TYPE "FRK_Document_D002"
VERSION : 0.1
   STRUCT
      SchemaVersion { ExternalAccessible := 'False'; ExternalVisible := 'False'; ExternalWritable := 'False'} : UInt;
      Scope { ExternalAccessible := 'False'; ExternalVisible := 'False'; ExternalWritable := 'False'} : String[80];
      Kind { ExternalAccessible := 'False'; ExternalVisible := 'False'; ExternalWritable := 'False'} : DInt;
      ModelCode { ExternalAccessible := 'False'; ExternalVisible := 'False'; ExternalWritable := 'False'} : String[64];
      ActiveModel { ExternalAccessible := 'False'; ExternalVisible := 'False'; ExternalWritable := 'False'} : String[64];
      Count { ExternalAccessible := 'False'; ExternalVisible := 'False'; ExternalWritable := 'False'} : Int;
      Rows { ExternalAccessible := 'False'; ExternalVisible := 'False'; ExternalWritable := 'False'} : Array[1..24] of "FRK_ConfigSlot";
   END_STRUCT;

END_TYPE

